(* IEC 61131-3 sources: trust-platform/crates/trust-runtime/tests/fixtures/plcopen_motion/single_axis_negative_group_label/src, 1 file *)

(* ---- tests.st ---- *)
TEST_PROGRAM plcopen_motion_single_axis_negative_group_label
VAR
    WrongAxisStatus : MC_AXIS_STATUS;
END_VAR

WrongAxisStatus := MC_AXIS_STATUS#GroupStandby;
END_TEST_PROGRAM
